Fanuc KAREL source: kb00155.KL

PROGRAM KB00155
%STACKSIZE=65535
%PRIORITY=65535
%NOLOCKGROUP
VAR
P1 : STRING[80]
P2 : INTEGER
BEGIN
P1='A'
P2=1
SAVE_DRAM(P1,P2)
END KB00155
